// TIA Portal V21 export
DATA_BLOCK "Controll_horizontale Achse_DB"   // DB5
// stored: InstanceOfName Controll_horizontale Achse, InstanceOfType FB
"Controll_horizontale Achse"
   // VAR_INPUT
   //    ModePos : Int;
   //    EnableAxis : Bool;
   //    IntermediateStop : Bool;
   //    AckError : Bool;
   //    ExecuteMode : Bool;
   //    Jog1 : Bool;
   //    Jog2 : Bool;
   //    Negative : Bool;
   //    Positive : Bool;
   //    Position : LReal;
   //    Velocity : LReal;
   // END_VAR
   // VAR_OUTPUT
   //    AxisEnabled : Bool;
   //    AxisPosOk : Bool;
   //    AxisRef : Bool;
   //    AxisError : Bool;
   //    Error : Bool;
   //    ActVelocity : LReal;
   //    ActPosition : LReal;
   // END_VAR
   // VAR
   //    Enable_XYMovement : Bool;
   //    AxisPos_max { ExternalAccessible := 'False'; ExternalVisible := 'False'; ExternalWritable := 'False'} : LReal;
   //    AxisPos_min { ExternalAccessible := 'False'; ExternalVisible := 'False'; ExternalWritable := 'False'} : LReal;
   // END_VAR
BEGIN
END_DATA_BLOCK
